(* IEC 61131-3 sources: plsim-chem/PLC, 4 files *)

(* ---- GVL_Sim.st ---- *)
// ---- GVL_Sim ----
{attribute 'qualified_only'}
VAR_GLOBAL
    P101_RunCmd : BOOL;  // P101.RunCmd: PLC writes (command)
    P101_SpeedSP : REAL;  // P101.SpeedSP: PLC writes (command)
    P101_ResetCmd : BOOL;  // P101.ResetCmd: PLC writes (command)
    P101_RunningFb : BOOL;  // P101.RunningFb: PLC reads (measurement/feedback)
    P101_Fault : BOOL;  // P101.Fault: PLC reads (measurement/feedback)
    P101_Speed : REAL;  // P101.Speed: PLC reads (measurement/feedback)
    P101_Current : REAL;  // P101.Current: PLC reads (measurement/feedback)
    P101_WindingTemp : REAL;  // P101.WindingTemp: PLC reads (measurement/feedback)
    P101_Voltage : REAL;  // P101.Voltage: PLC reads (measurement/feedback)
    P101_Vibration : REAL;  // P101.Vibration: PLC reads (measurement/feedback)
    P102_RunCmd : BOOL;  // P102.RunCmd: PLC writes (command)
    P102_SpeedSP : REAL;  // P102.SpeedSP: PLC writes (command)
    P102_ResetCmd : BOOL;  // P102.ResetCmd: PLC writes (command)
    P102_RunningFb : BOOL;  // P102.RunningFb: PLC reads (measurement/feedback)
    P102_Fault : BOOL;  // P102.Fault: PLC reads (measurement/feedback)
    P102_Speed : REAL;  // P102.Speed: PLC reads (measurement/feedback)
    P102_Current : REAL;  // P102.Current: PLC reads (measurement/feedback)
    P102_WindingTemp : REAL;  // P102.WindingTemp: PLC reads (measurement/feedback)
    P102_Voltage : REAL;  // P102.Voltage: PLC reads (measurement/feedback)
    P102_Vibration : REAL;  // P102.Vibration: PLC reads (measurement/feedback)
    P103_RunCmd : BOOL;  // P103.RunCmd: PLC writes (command)
    P103_SpeedSP : REAL;  // P103.SpeedSP: PLC writes (command)
    P103_ResetCmd : BOOL;  // P103.ResetCmd: PLC writes (command)
    P103_RunningFb : BOOL;  // P103.RunningFb: PLC reads (measurement/feedback)
    P103_Fault : BOOL;  // P103.Fault: PLC reads (measurement/feedback)
    P103_Speed : REAL;  // P103.Speed: PLC reads (measurement/feedback)
    P103_Current : REAL;  // P103.Current: PLC reads (measurement/feedback)
    P103_WindingTemp : REAL;  // P103.WindingTemp: PLC reads (measurement/feedback)
    P103_Voltage : REAL;  // P103.Voltage: PLC reads (measurement/feedback)
    P103_Vibration : REAL;  // P103.Vibration: PLC reads (measurement/feedback)
    XV101_OpenCmd : BOOL;  // XV101.OpenCmd: PLC writes (command)
    XV101_PositionSP : REAL;  // XV101.PositionSP: PLC writes (command)
    XV101_OpenFb : BOOL;  // XV101.OpenFb: PLC reads (measurement/feedback)
    XV101_ClosedFb : BOOL;  // XV101.ClosedFb: PLC reads (measurement/feedback)
    XV101_Position : REAL;  // XV101.Position: PLC reads (measurement/feedback)
    XV102_OpenCmd : BOOL;  // XV102.OpenCmd: PLC writes (command)
    XV102_PositionSP : REAL;  // XV102.PositionSP: PLC writes (command)
    XV102_OpenFb : BOOL;  // XV102.OpenFb: PLC reads (measurement/feedback)
    XV102_ClosedFb : BOOL;  // XV102.ClosedFb: PLC reads (measurement/feedback)
    XV102_Position : REAL;  // XV102.Position: PLC reads (measurement/feedback)
    XV103_OpenCmd : BOOL;  // XV103.OpenCmd: PLC writes (command)
    XV103_PositionSP : REAL;  // XV103.PositionSP: PLC writes (command)
    XV103_OpenFb : BOOL;  // XV103.OpenFb: PLC reads (measurement/feedback)
    XV103_ClosedFb : BOOL;  // XV103.ClosedFb: PLC reads (measurement/feedback)
    XV103_Position : REAL;  // XV103.Position: PLC reads (measurement/feedback)
    XV111_OpenCmd : BOOL;  // XV111.OpenCmd: PLC writes (command)
    XV111_PositionSP : REAL;  // XV111.PositionSP: PLC writes (command)
    XV111_OpenFb : BOOL;  // XV111.OpenFb: PLC reads (measurement/feedback)
    XV111_ClosedFb : BOOL;  // XV111.ClosedFb: PLC reads (measurement/feedback)
    XV111_Position : REAL;  // XV111.Position: PLC reads (measurement/feedback)
    XV112_OpenCmd : BOOL;  // XV112.OpenCmd: PLC writes (command)
    XV112_PositionSP : REAL;  // XV112.PositionSP: PLC writes (command)
    XV112_OpenFb : BOOL;  // XV112.OpenFb: PLC reads (measurement/feedback)
    XV112_ClosedFb : BOOL;  // XV112.ClosedFb: PLC reads (measurement/feedback)
    XV112_Position : REAL;  // XV112.Position: PLC reads (measurement/feedback)
    XV113_OpenCmd : BOOL;  // XV113.OpenCmd: PLC writes (command)
    XV113_PositionSP : REAL;  // XV113.PositionSP: PLC writes (command)
    XV113_OpenFb : BOOL;  // XV113.OpenFb: PLC reads (measurement/feedback)
    XV113_ClosedFb : BOOL;  // XV113.ClosedFb: PLC reads (measurement/feedback)
    XV113_Position : REAL;  // XV113.Position: PLC reads (measurement/feedback)
    XV201_OpenCmd : BOOL;  // XV201.OpenCmd: PLC writes (command)
    XV201_PositionSP : REAL;  // XV201.PositionSP: PLC writes (command)
    XV201_OpenFb : BOOL;  // XV201.OpenFb: PLC reads (measurement/feedback)
    XV201_ClosedFb : BOOL;  // XV201.ClosedFb: PLC reads (measurement/feedback)
    XV201_Position : REAL;  // XV201.Position: PLC reads (measurement/feedback)
    XV210_OpenCmd : BOOL;  // XV210.OpenCmd: PLC writes (command)
    XV210_PositionSP : REAL;  // XV210.PositionSP: PLC writes (command)
    XV210_OpenFb : BOOL;  // XV210.OpenFb: PLC reads (measurement/feedback)
    XV210_ClosedFb : BOOL;  // XV210.ClosedFb: PLC reads (measurement/feedback)
    XV210_Position : REAL;  // XV210.Position: PLC reads (measurement/feedback)
    AT201_Value : REAL;  // AT201.Value: PLC reads (measurement/feedback)
    AT201_Raw : INT;  // AT201.Raw: PLC reads (measurement/feedback)
    FT101_Value : REAL;  // FT101.Value: PLC reads (measurement/feedback)
    FT101_Raw : INT;  // FT101.Raw: PLC reads (measurement/feedback)
    FT102_Value : REAL;  // FT102.Value: PLC reads (measurement/feedback)
    FT102_Raw : INT;  // FT102.Raw: PLC reads (measurement/feedback)
    FT103_Value : REAL;  // FT103.Value: PLC reads (measurement/feedback)
    FT103_Raw : INT;  // FT103.Raw: PLC reads (measurement/feedback)
    FT201_Value : REAL;  // FT201.Value: PLC reads (measurement/feedback)
    FT201_Raw : INT;  // FT201.Raw: PLC reads (measurement/feedback)
    LT101_Value : REAL;  // LT101.Value: PLC reads (measurement/feedback)
    LT101_Raw : INT;  // LT101.Raw: PLC reads (measurement/feedback)
    LT102_Value : REAL;  // LT102.Value: PLC reads (measurement/feedback)
    LT102_Raw : INT;  // LT102.Raw: PLC reads (measurement/feedback)
    LT103_Value : REAL;  // LT103.Value: PLC reads (measurement/feedback)
    LT103_Raw : INT;  // LT103.Raw: PLC reads (measurement/feedback)
    LT201_Value : REAL;  // LT201.Value: PLC reads (measurement/feedback)
    LT201_Raw : INT;  // LT201.Raw: PLC reads (measurement/feedback)
    PDT111_Value : REAL;  // PDT111.Value: PLC reads (measurement/feedback)
    PDT111_Raw : INT;  // PDT111.Raw: PLC reads (measurement/feedback)
    PT101_Value : REAL;  // PT101.Value: PLC reads (measurement/feedback)
    PT101_Raw : INT;  // PT101.Raw: PLC reads (measurement/feedback)
    TT201_Value : REAL;  // TT201.Value: PLC reads (measurement/feedback)
    TT201_Raw : INT;  // TT201.Raw: PLC reads (measurement/feedback)
END_VAR

(* ---- GVL_Sim_demo.st ---- *)
// ---- GVL_Sim ----
{attribute 'qualified_only'}
VAR_GLOBAL
    C301_HeaterCmd : REAL;  // C301.HeaterCmd: PLC writes (command)
    C301_RefluxCmd : REAL;  // C301.RefluxCmd: PLC writes (command)
    C301_TopTemp : REAL;  // C301.TopTemp: PLC reads (measurement/feedback)
    C301_BottomTemp : REAL;  // C301.BottomTemp: PLC reads (measurement/feedback)
    C301_Boilup : REAL;  // C301.Boilup: PLC reads (measurement/feedback)
    C301_DrumLevel : REAL;  // C301.DrumLevel: PLC reads (measurement/feedback)
    C301_ColumnDp : REAL;  // C301.ColumnDp: PLC reads (measurement/feedback)
    C301_Flooding : BOOL;  // C301.Flooding: PLC reads (measurement/feedback)
    CP301_RunCmd : BOOL;  // CP301.RunCmd: PLC writes (command)
    CP301_SpeedSP : REAL;  // CP301.SpeedSP: PLC writes (command)
    CP301_ResetCmd : BOOL;  // CP301.ResetCmd: PLC writes (command)
    CP301_RunningFb : BOOL;  // CP301.RunningFb: PLC reads (measurement/feedback)
    CP301_Fault : BOOL;  // CP301.Fault: PLC reads (measurement/feedback)
    CP301_Surge : BOOL;  // CP301.Surge: PLC reads (measurement/feedback)
    CP301_Speed : REAL;  // CP301.Speed: PLC reads (measurement/feedback)
    CP301_Power : REAL;  // CP301.Power: PLC reads (measurement/feedback)
    CP301_DischargeTemp : REAL;  // CP301.DischargeTemp: PLC reads (measurement/feedback)
    CP301_Current : REAL;  // CP301.Current: PLC reads (measurement/feedback)
    CP301_WindingTemp : REAL;  // CP301.WindingTemp: PLC reads (measurement/feedback)
    CP301_Voltage : REAL;  // CP301.Voltage: PLC reads (measurement/feedback)
    CP301_Vibration : REAL;  // CP301.Vibration: PLC reads (measurement/feedback)
    EV301_HeaterCmd : REAL;  // EV301.HeaterCmd: PLC writes (command)
    EV301_CoolingCmd : REAL;  // EV301.CoolingCmd: PLC writes (command)
    EV301_EvapRate : REAL;  // EV301.EvapRate: PLC reads (measurement/feedback)
    GVV301_OpenCmd : BOOL;  // GVV301.OpenCmd: PLC writes (command)
    GVV301_PositionSP : REAL;  // GVV301.PositionSP: PLC writes (command)
    GVV301_OpenFb : BOOL;  // GVV301.OpenFb: PLC reads (measurement/feedback)
    GVV301_ClosedFb : BOOL;  // GVV301.ClosedFb: PLC reads (measurement/feedback)
    GVV301_Position : REAL;  // GVV301.Position: PLC reads (measurement/feedback)
    HX301_DutyCmd : REAL;  // HX301.DutyCmd: PLC writes (command)
    HX301_Duty : REAL;  // HX301.Duty: PLC reads (measurement/feedback)
    HX301_OutletTemp : REAL;  // HX301.OutletTemp: PLC reads (measurement/feedback)
    P301_RunCmd : BOOL;  // P301.RunCmd: PLC writes (command)
    P301_SpeedSP : REAL;  // P301.SpeedSP: PLC writes (command)
    P301_ResetCmd : BOOL;  // P301.ResetCmd: PLC writes (command)
    P301_RunningFb : BOOL;  // P301.RunningFb: PLC reads (measurement/feedback)
    P301_Fault : BOOL;  // P301.Fault: PLC reads (measurement/feedback)
    P301_Speed : REAL;  // P301.Speed: PLC reads (measurement/feedback)
    P301_Current : REAL;  // P301.Current: PLC reads (measurement/feedback)
    P301_WindingTemp : REAL;  // P301.WindingTemp: PLC reads (measurement/feedback)
    P301_Voltage : REAL;  // P301.Voltage: PLC reads (measurement/feedback)
    P301_Vibration : REAL;  // P301.Vibration: PLC reads (measurement/feedback)
    P302_RunCmd : BOOL;  // P302.RunCmd: PLC writes (command)
    P302_SpeedSP : REAL;  // P302.SpeedSP: PLC writes (command)
    P302_ResetCmd : BOOL;  // P302.ResetCmd: PLC writes (command)
    P302_RunningFb : BOOL;  // P302.RunningFb: PLC reads (measurement/feedback)
    P302_Fault : BOOL;  // P302.Fault: PLC reads (measurement/feedback)
    P302_Speed : REAL;  // P302.Speed: PLC reads (measurement/feedback)
    P302_Current : REAL;  // P302.Current: PLC reads (measurement/feedback)
    P302_WindingTemp : REAL;  // P302.WindingTemp: PLC reads (measurement/feedback)
    P302_Voltage : REAL;  // P302.Voltage: PLC reads (measurement/feedback)
    P302_Vibration : REAL;  // P302.Vibration: PLC reads (measurement/feedback)
    P303_RunCmd : BOOL;  // P303.RunCmd: PLC writes (command)
    P303_SpeedSP : REAL;  // P303.SpeedSP: PLC writes (command)
    P303_ResetCmd : BOOL;  // P303.ResetCmd: PLC writes (command)
    P303_RunningFb : BOOL;  // P303.RunningFb: PLC reads (measurement/feedback)
    P303_Fault : BOOL;  // P303.Fault: PLC reads (measurement/feedback)
    P303_Speed : REAL;  // P303.Speed: PLC reads (measurement/feedback)
    P303_Current : REAL;  // P303.Current: PLC reads (measurement/feedback)
    P303_WindingTemp : REAL;  // P303.WindingTemp: PLC reads (measurement/feedback)
    P303_Voltage : REAL;  // P303.Voltage: PLC reads (measurement/feedback)
    P303_Vibration : REAL;  // P303.Vibration: PLC reads (measurement/feedback)
    XV301_OpenCmd : BOOL;  // XV301.OpenCmd: PLC writes (command)
    XV301_PositionSP : REAL;  // XV301.PositionSP: PLC writes (command)
    XV301_OpenFb : BOOL;  // XV301.OpenFb: PLC reads (measurement/feedback)
    XV301_ClosedFb : BOOL;  // XV301.ClosedFb: PLC reads (measurement/feedback)
    XV301_Position : REAL;  // XV301.Position: PLC reads (measurement/feedback)
    XV302_OpenCmd : BOOL;  // XV302.OpenCmd: PLC writes (command)
    XV302_PositionSP : REAL;  // XV302.PositionSP: PLC writes (command)
    XV302_OpenFb : BOOL;  // XV302.OpenFb: PLC reads (measurement/feedback)
    XV302_ClosedFb : BOOL;  // XV302.ClosedFb: PLC reads (measurement/feedback)
    XV302_Position : REAL;  // XV302.Position: PLC reads (measurement/feedback)
    AT302_Value : REAL;  // AT302.Value: PLC reads (measurement/feedback)
    AT302_Raw : INT;  // AT302.Raw: PLC reads (measurement/feedback)
    FT301_Value : REAL;  // FT301.Value: PLC reads (measurement/feedback)
    FT301_Raw : INT;  // FT301.Raw: PLC reads (measurement/feedback)
    FT302_Value : REAL;  // FT302.Value: PLC reads (measurement/feedback)
    FT302_Raw : INT;  // FT302.Raw: PLC reads (measurement/feedback)
    LT301_Value : REAL;  // LT301.Value: PLC reads (measurement/feedback)
    LT301_Raw : INT;  // LT301.Raw: PLC reads (measurement/feedback)
    LT302_Value : REAL;  // LT302.Value: PLC reads (measurement/feedback)
    LT302_Raw : INT;  // LT302.Raw: PLC reads (measurement/feedback)
    LT303_Value : REAL;  // LT303.Value: PLC reads (measurement/feedback)
    LT303_Raw : INT;  // LT303.Raw: PLC reads (measurement/feedback)
    PDT301_Value : REAL;  // PDT301.Value: PLC reads (measurement/feedback)
    PDT301_Raw : INT;  // PDT301.Raw: PLC reads (measurement/feedback)
    PT301_Value : REAL;  // PT301.Value: PLC reads (measurement/feedback)
    PT301_Raw : INT;  // PT301.Raw: PLC reads (measurement/feedback)
    TT301_Value : REAL;  // TT301.Value: PLC reads (measurement/feedback)
    TT301_Raw : INT;  // TT301.Raw: PLC reads (measurement/feedback)
    TT302_Value : REAL;  // TT302.Value: PLC reads (measurement/feedback)
    TT302_Raw : INT;  // TT302.Raw: PLC reads (measurement/feedback)
    TT303_Value : REAL;  // TT303.Value: PLC reads (measurement/feedback)
    TT303_Raw : INT;  // TT303.Raw: PLC reads (measurement/feedback)
END_VAR

(* ---- GVL_Sim_training.st ---- *)
// ---- GVL_Sim ----
{attribute 'qualified_only'}
VAR_GLOBAL
    P401_RunCmd : BOOL;  // P401.RunCmd: PLC writes (command)
    P401_SpeedSP : REAL;  // P401.SpeedSP: PLC writes (command)
    P401_ResetCmd : BOOL;  // P401.ResetCmd: PLC writes (command)
    P401_RunningFb : BOOL;  // P401.RunningFb: PLC reads (measurement/feedback)
    P401_Fault : BOOL;  // P401.Fault: PLC reads (measurement/feedback)
    P401_Speed : REAL;  // P401.Speed: PLC reads (measurement/feedback)
    P401_Current : REAL;  // P401.Current: PLC reads (measurement/feedback)
    P401_WindingTemp : REAL;  // P401.WindingTemp: PLC reads (measurement/feedback)
    P401_Voltage : REAL;  // P401.Voltage: PLC reads (measurement/feedback)
    P401_Vibration : REAL;  // P401.Vibration: PLC reads (measurement/feedback)
    P402_RunCmd : BOOL;  // P402.RunCmd: PLC writes (command)
    P402_SpeedSP : REAL;  // P402.SpeedSP: PLC writes (command)
    P402_ResetCmd : BOOL;  // P402.ResetCmd: PLC writes (command)
    P402_RunningFb : BOOL;  // P402.RunningFb: PLC reads (measurement/feedback)
    P402_Fault : BOOL;  // P402.Fault: PLC reads (measurement/feedback)
    P402_Speed : REAL;  // P402.Speed: PLC reads (measurement/feedback)
    P402_Current : REAL;  // P402.Current: PLC reads (measurement/feedback)
    P402_WindingTemp : REAL;  // P402.WindingTemp: PLC reads (measurement/feedback)
    P402_Voltage : REAL;  // P402.Voltage: PLC reads (measurement/feedback)
    P402_Vibration : REAL;  // P402.Vibration: PLC reads (measurement/feedback)
    UV401_OpenCmd : BOOL;  // UV401.OpenCmd: PLC writes (command)
    UV401_PositionSP : REAL;  // UV401.PositionSP: PLC writes (command)
    UV401_OpenFb : BOOL;  // UV401.OpenFb: PLC reads (measurement/feedback)
    UV401_ClosedFb : BOOL;  // UV401.ClosedFb: PLC reads (measurement/feedback)
    UV401_Position : REAL;  // UV401.Position: PLC reads (measurement/feedback)
    UV402_OpenCmd : BOOL;  // UV402.OpenCmd: PLC writes (command)
    UV402_PositionSP : REAL;  // UV402.PositionSP: PLC writes (command)
    UV402_OpenFb : BOOL;  // UV402.OpenFb: PLC reads (measurement/feedback)
    UV402_ClosedFb : BOOL;  // UV402.ClosedFb: PLC reads (measurement/feedback)
    UV402_Position : REAL;  // UV402.Position: PLC reads (measurement/feedback)
    XV402_OpenCmd : BOOL;  // XV402.OpenCmd: PLC writes (command)
    XV402_PositionSP : REAL;  // XV402.PositionSP: PLC writes (command)
    XV402_OpenFb : BOOL;  // XV402.OpenFb: PLC reads (measurement/feedback)
    XV402_ClosedFb : BOOL;  // XV402.ClosedFb: PLC reads (measurement/feedback)
    XV402_Position : REAL;  // XV402.Position: PLC reads (measurement/feedback)
    XV404_OpenCmd : BOOL;  // XV404.OpenCmd: PLC writes (command)
    XV404_PositionSP : REAL;  // XV404.PositionSP: PLC writes (command)
    XV404_OpenFb : BOOL;  // XV404.OpenFb: PLC reads (measurement/feedback)
    XV404_ClosedFb : BOOL;  // XV404.ClosedFb: PLC reads (measurement/feedback)
    XV404_Position : REAL;  // XV404.Position: PLC reads (measurement/feedback)
    AT401_Value : REAL;  // AT401.Value: PLC reads (measurement/feedback)
    AT401_Raw : INT;  // AT401.Raw: PLC reads (measurement/feedback)
    AT402_Value : REAL;  // AT402.Value: PLC reads (measurement/feedback)
    AT402_Raw : INT;  // AT402.Raw: PLC reads (measurement/feedback)
    FT401_Value : REAL;  // FT401.Value: PLC reads (measurement/feedback)
    FT401_Raw : INT;  // FT401.Raw: PLC reads (measurement/feedback)
    FT402_Value : REAL;  // FT402.Value: PLC reads (measurement/feedback)
    FT402_Raw : INT;  // FT402.Raw: PLC reads (measurement/feedback)
    LT401_Value : REAL;  // LT401.Value: PLC reads (measurement/feedback)
    LT401_Raw : INT;  // LT401.Raw: PLC reads (measurement/feedback)
    LT402_Value : REAL;  // LT402.Value: PLC reads (measurement/feedback)
    LT402_Raw : INT;  // LT402.Raw: PLC reads (measurement/feedback)
    PDT402_Value : REAL;  // PDT402.Value: PLC reads (measurement/feedback)
    PDT402_Raw : INT;  // PDT402.Raw: PLC reads (measurement/feedback)
    PDT404_Value : REAL;  // PDT404.Value: PLC reads (measurement/feedback)
    PDT404_Raw : INT;  // PDT404.Raw: PLC reads (measurement/feedback)
    PT401_Value : REAL;  // PT401.Value: PLC reads (measurement/feedback)
    PT401_Raw : INT;  // PT401.Raw: PLC reads (measurement/feedback)
    PT402_Value : REAL;  // PT402.Value: PLC reads (measurement/feedback)
    PT402_Raw : INT;  // PT402.Raw: PLC reads (measurement/feedback)
    TT401_Value : REAL;  // TT401.Value: PLC reads (measurement/feedback)
    TT401_Raw : INT;  // TT401.Raw: PLC reads (measurement/feedback)
    TT402_Value : REAL;  // TT402.Value: PLC reads (measurement/feedback)
    TT402_Raw : INT;  // TT402.Raw: PLC reads (measurement/feedback)
END_VAR

(* ---- MAIN_example.st ---- *)
// =====================================================================
// MAIN_example.st : starter PLC program for the test plant
// Paste into a TwinCAT PLC program called MAIN. Needs the GVL_Sim variables from GVL_Sim.st.
//
// What it does
//  - Keeps each feed tank between 70 % and 90 % by opening its inlet valve (hysteresis)
//  - Pumps feed from the tanks to the reactor while the reactor is below 70 %
//  - A pump only runs when its tank is not empty and its outlet valve is confirmed open
//  - Cooling water valve follows the reactor temperature (proportional control)
//  - Latching safety trip on high temperature or high reactor level
//
// Set bRun to TRUE (online, or from the HMI) to start. Set bReset to TRUE to clear a trip or a pump fault.
// Variables that the simulation writes (..Value, ..Raw, ..OpenFb, ..ClosedFb, ..RunningFb, ..Fault, ..Position, ..Speed)
// must only be read here. Variables ending in ..OpenCmd, ..RunCmd, ..ResetCmd, ..SpeedSP, ..PositionSP are yours to write.
// =====================================================================

PROGRAM MAIN
VAR
    bRun            : BOOL;             // operator: start the sequence
    bReset          : BOOL;             // operator: reset trip and pump faults
    bTrip           : BOOL;             // latched safety trip
    bTransfer       : BOOL;             // feed transfer to the reactor is allowed
    bFill1          : BOOL;
    bFill2          : BOOL;
    bFill3          : BOOL;

    rTempSP         : REAL := 40.0;     // reactor temperature setpoint, C
    rTempTrip       : REAL := 70.0;     // trip above this temperature, C
    rLevelMax       : REAL := 70.0;     // stop transfer at this reactor level, %
    rLevelTrip      : REAL := 90.0;     // trip at this reactor level, %
    rCoolingGain    : REAL := 6.0;      // % valve opening per C above setpoint
    rCooling        : REAL;
END_VAR

// ---- Safety trip ----------------------------------------------------
IF GVL_Sim.TT201_Value > rTempTrip OR GVL_Sim.LT201_Value > rLevelTrip THEN
    bTrip := TRUE;
END_IF
IF bReset AND GVL_Sim.TT201_Value < rTempSP + 10.0 AND GVL_Sim.LT201_Value < rLevelMax THEN
    bTrip := FALSE;
END_IF

// ---- Feed tank filling (hysteresis) ---------------------------------
IF GVL_Sim.LT101_Value < 70.0 THEN bFill1 := TRUE; ELSIF GVL_Sim.LT101_Value > 90.0 THEN bFill1 := FALSE; END_IF
IF GVL_Sim.LT102_Value < 70.0 THEN bFill2 := TRUE; ELSIF GVL_Sim.LT102_Value > 90.0 THEN bFill2 := FALSE; END_IF
IF GVL_Sim.LT103_Value < 70.0 THEN bFill3 := TRUE; ELSIF GVL_Sim.LT103_Value > 90.0 THEN bFill3 := FALSE; END_IF

GVL_Sim.XV101_OpenCmd := bRun AND NOT bTrip AND bFill1;
GVL_Sim.XV102_OpenCmd := bRun AND NOT bTrip AND bFill2;
GVL_Sim.XV103_OpenCmd := bRun AND NOT bTrip AND bFill3;

// ---- Transfer to the reactor (hysteresis on reactor level) ----------
IF NOT bRun OR bTrip OR GVL_Sim.LT201_Value >= rLevelMax THEN
    bTransfer := FALSE;
ELSIF GVL_Sim.LT201_Value <= rLevelMax - 10.0 THEN
    bTransfer := TRUE;
END_IF

GVL_Sim.XV111_OpenCmd := bTransfer;
GVL_Sim.XV112_OpenCmd := bTransfer;
GVL_Sim.XV113_OpenCmd := bTransfer;

GVL_Sim.P101_RunCmd := bTransfer AND GVL_Sim.XV111_OpenFb AND GVL_Sim.LT101_Value > 10.0 AND NOT GVL_Sim.P101_Fault;
GVL_Sim.P102_RunCmd := bTransfer AND GVL_Sim.XV112_OpenFb AND GVL_Sim.LT102_Value > 10.0 AND NOT GVL_Sim.P102_Fault;
GVL_Sim.P103_RunCmd := bTransfer AND GVL_Sim.XV113_OpenFb AND GVL_Sim.LT103_Value > 10.0 AND NOT GVL_Sim.P103_Fault;
GVL_Sim.P103_SpeedSP := 40.0;       // water pump is variable speed

GVL_Sim.P101_ResetCmd := bReset;
GVL_Sim.P102_ResetCmd := bReset;
GVL_Sim.P103_ResetCmd := bReset;

// ---- Reactor cooling (proportional) and outlet -----------------------
rCooling := 20.0 + rCoolingGain * (GVL_Sim.TT201_Value - rTempSP);
GVL_Sim.XV210_PositionSP := LIMIT(0.0, rCooling, 100.0);

IF bRun AND NOT bTrip AND GVL_Sim.LT201_Value > 30.0 THEN
    GVL_Sim.XV201_PositionSP := 60.0;
ELSE
    GVL_Sim.XV201_PositionSP := 0.0;
END_IF
